Fanuc KAREL source: KT00287.KL

PROGRAM KT00287
%NOLOCKGROUP
VAR
  P1: JOINTPOS
  P2: POSITION
  OUT: BOOLEAN
BEGIN
  OUT = P1 = P2
END KT00287
